FUNCTION_BLOCK HYST_SM
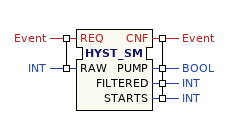
  EVENT_INPUT
    REQ WITH RAW;
  END_EVENT
  EVENT_OUTPUT
    CNF WITH PUMP, FILTERED, STARTS;
  END_EVENT
  VAR_INPUT
    RAW : INT;
  END_VAR
  VAR_OUTPUT
    PUMP : BOOL;
    FILTERED : INT;
    STARTS : INT;
  END_VAR
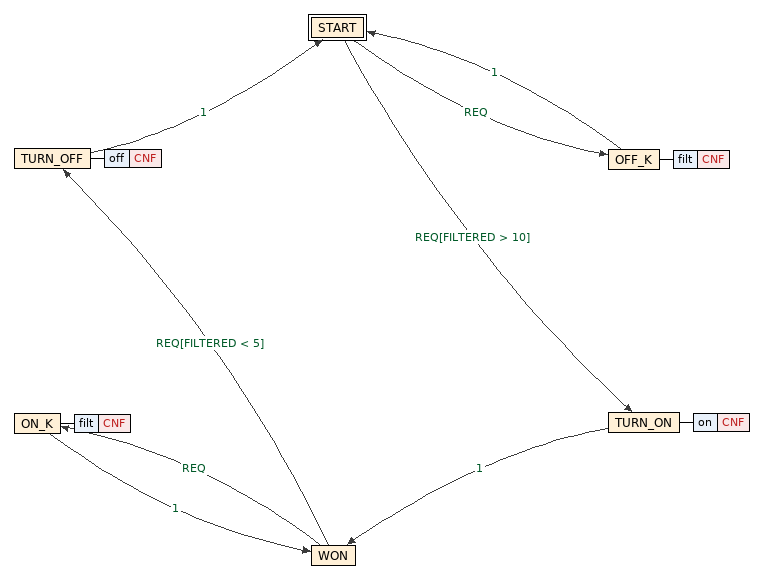
  EC_STATES
    START;
    OFF_K : filt -> CNF;
    TURN_ON : on -> CNF;
    WON;
    ON_K : filt -> CNF;
    TURN_OFF : off -> CNF;
  END_STATES
  EC_TRANSITIONS
    START TO TURN_ON := REQ[FILTERED > 10];
    START TO OFF_K := REQ;
    OFF_K TO START := 1;
    TURN_ON TO WON := 1;
    WON TO TURN_OFF := REQ[FILTERED < 5];
    WON TO ON_K := REQ;
    ON_K TO WON := 1;
    TURN_OFF TO START := 1;
  END_TRANSITIONS
  ALGORITHM filt IN ST:
FILTERED := (FILTERED + RAW) / 2;
  END_ALGORITHM
  ALGORITHM on IN ST:
PUMP := TRUE;
STARTS := STARTS + 1;
FILTERED := (FILTERED + RAW) / 2;
  END_ALGORITHM
  ALGORITHM off IN ST:
PUMP := FALSE;
FILTERED := (FILTERED + RAW) / 2;
  END_ALGORITHM
END_FUNCTION_BLOCK
